// TwinCAT 3 PLC project PLC
// ProgramVersion: 3.1.4026.27
// CompilerDefines: VISU_USEPROPERTYINFO
// libraries:
//   Tc2_Standard, * (Beckhoff Automation GmbH)
//   Tc2_System, * (Beckhoff Automation GmbH)
//   Tc2_Utilities, * (Beckhoff Automation GmbH)
//   Tc3_DynamicMemory, * (Beckhoff Automation GmbH)
//   VisuDialogs, * (System)
//   VisuSymbols, 4.5.0.0 (System)
// project tree:
//   / GlobalTextList.TcGTLO, PlcTask.TcTTO, Visualization Manager.TcVMO (not stored)
//   POUs/ FB_Dynamic.TcPOU, MAIN.TcPOU, monoInstance.TcPOU, multiInstances.TcPOU
//   VISUs/ Visualization.TcVIS
// real-time tasks:
//   TASK PlcTask: cycle T#10ms, priority 20, ADS port 350

CONFIGURATION PLC
    RESOURCE PLC ON TwinCAT3
        TASK PlcTask(INTERVAL := T#10ms, PRIORITY := 20);
        PROGRAM MAIN WITH PlcTask : MAIN;
    END_RESOURCE
END_CONFIGURATION

// ---- POUs/MAIN.TcPOU
PROGRAM MAIN
VAR
(*
+--------------------------------------------------------------------------+
| PROGRAMME DE TEST - CREATION DYNAMIQUE (__NEW / __DELETE)                |
| TwinCAT 3 - IEC 61131-3 - Structured Text                                |
+--------------------------------------------------------------------------+
|                                                                          |
| Projet d'exemple TwinCAT 3 illustrant la creation et la destruction      |
| dynamiques d'instances de bloc fonction (FB) pendant l'execution du      |
| PLC, avec les operateurs __NEW et __DELETE.                              |
|                                                                          |
+--------------------------------------------------------------------------+
| monoInstance                                                             |
|   -> Creer / detruire une seule instance de FB_Dynamic                   |
+--------------------------------------------------------------------------+
| multiInstances                                                           |
|   -> Gerer un nombre dynamique d'instances (de 0 a cMaxInstances),       |
|      ajustable en ligne, avec suivi de la memoire du router              |
+--------------------------------------------------------------------------+
*)
END_VAR

//monoInstance();
multiInstances();

END_PROGRAM

// ---- POUs/multiInstances.TcPOU
PROGRAM multiInstances
VAR CONSTANT
    cMaxInstances : UINT := 1000;      // passer à 100, puis 1000 pour tester les limites
END_VAR
VAR
    // Tableau de pointeurs (aucune instance n'est créée statiquement)
    aFB            : ARRAY[1..cMaxInstances] OF POINTER TO FB_Dynamic;
    aResult        : ARRAY[1..cMaxInstances] OF INT;

    // Commande
    nTarget        : UINT := 10;     // nombre d'instances souhaité (modifiable en ligne)
    nMaxOpsPerCycle: UINT := 50;     // limite de __NEW/__DELETE par cycle
    nIncrease      : INT := 5;

    // Diagnostic
    nActive        : UINT;           // instances actuellement créées
    nNewFailed     : UDINT;          // nombre d'échecs de __NEW
    bAllocError    : BOOL;

    // Variables locales de travail
    i              : UINT;
    nOps           : UINT;

    // Surveillance du router (ton code existant)
    fbGetRouterStatusInfo : FB_GetRouterStatusInfo;
    TonGetRouterStatus    : TON;
    bError                : BOOL;
    nErrorID              : UDINT;
    stTcRouterStatusInfo  : Tc2_Utilities.ST_TcRouterStatusInfo;
	nUsage: REAL;
	bInc: BOOL;
	bDec: BOOL;
END_VAR

// --- 1. Ajustement du nombre d'instances vers nTarget ---
nTarget := LIMIT(0, nTarget, cMaxInstances);
nOps    := 0;

FOR i := 1 TO cMaxInstances DO
    IF nOps >= nMaxOpsPerCycle THEN
        EXIT;                              // on étale la charge sur plusieurs cycles
    END_IF

    IF i <= nTarget THEN
        // Instance souhaitée : on la crée si elle n'existe pas
        IF aFB[i] = 0 THEN
            aFB[i] := __NEW(FB_Dynamic);
            nOps := nOps + 1;
            IF aFB[i] = 0 THEN             // __NEW renvoie 0 si plus de mémoire
                nNewFailed  := nNewFailed + 1;
                bAllocError := TRUE;
                EXIT;
            END_IF
        END_IF
    ELSE
        // Instance en trop : on la détruit
        IF aFB[i] <> 0 THEN
            __DELETE(aFB[i]);
            aFB[i] := 0;                   // indispensable
            nOps := nOps + 1;
        END_IF
    END_IF
END_FOR

// --- 2. Appel cyclique des instances existantes ---
nActive := 0;
FOR i := 1 TO cMaxInstances DO
    IF aFB[i] <> 0 THEN
        aResult[i] := aFB[i]^.Increase(nCountStep := nIncrease);
        nActive    := nActive + 1;
    END_IF
END_FOR

// --- 3. Surveillance du router (inchangé) ---
fbGetRouterStatusInfo(
    sNetId   := '',
    bExecute := NOT TonGetRouterStatus.Q,
    tTimeout := DEFAULT_ADS_TIMEOUT,
    bBusy    => ,
    bError   => bError,
    nErrID   => nErrorID,
    info     => stTcRouterStatusInfo);

TonGetRouterStatus(IN := NOT fbGetRouterStatusInfo.bBusy, PT := T#1S);

IF stTcRouterStatusInfo.maxMem >0 THEN
nUsage:=(TO_REAL(stTcRouterStatusInfo.maxMem-stTcRouterStatusInfo.maxMemAvail)/TO_REAL(stTcRouterStatusInfo.maxMem))*100.0;
END_IF

IF bInc AND nTarget<cMaxInstances THEN
	nTarget:=nTarget+1;
	bInc:=FALSE;
END_IF

IF bDec  AND nTarget>1 THEN
	nTarget:=nTarget-1;
	bDec:=FALSE;
END_IF

END_PROGRAM

// ---- POUs/FB_Dynamic.TcPOU
{attribute 'enable_dynamic_creation'}
FUNCTION_BLOCK FB_Dynamic
VAR
    nCounts : INT;
END_VAR

METHOD Increase : INT
VAR_INPUT
	nCountStep :INT;
END_VAR
nCounts := nCounts + nCountStep;
Increase := nCounts;
END_METHOD

END_FUNCTION_BLOCK

// ---- POUs/monoInstance.TcPOU
PROGRAM monoInstance
VAR
	pFB       : POINTER TO FB_Dynamic;
    nResult   : INT;
    nIncrease : INT := 5;
    bNew      : BOOL := TRUE;
    bDelete   : BOOL;
	
	fbGetRouterStatusInfo:FB_GetRouterStatusInfo;
	TonGetRouterStatus:TON;
	bError: BOOL;
	nErrorID: UDINT;
	stTcRouterStatusInfo: Tc2_Utilities.ST_TcRouterStatusInfo;
END_VAR

IF bNew AND (pFB = 0) THEN
    pFB := __NEW(FB_Dynamic);
    bNew := FALSE;
END_IF

IF (pFB <> 0) THEN
    nResult := pFB^.Increase(nCountStep := nIncrease);
END_IF

IF bDelete THEN
    __DELETE(pFB);
    bDelete := FALSE;
END_IF


fbGetRouterStatusInfo(
	sNetId:= '', 
	bExecute:= NOT TonGetRouterStatus.Q, 
	tTimeout:= DEFAULT_ADS_TIMEOUT, 
	bBusy=> , 
	bError=> bError, 
	nErrID=> nErrorID, 
	info=> stTcRouterStatusInfo);

IF stTcRouterStatusInfo.maxMem >0 THEN
	TonGetRouterStatus(IN:= NOT fbGetRouterStatusInfo.bBusy, PT:=T#1S , Q=> , ET=> );
END_IF

END_PROGRAM

// ---- GlobalTextList.TcGTLO
TEXTLIST GlobalTextList
  77 = '+'
  247 = '-'
  9 = 'nb Instances %d'
  278 = 'nb Instances: %d'
  284 = 'nb Target: %d'
  238 = 'Usage : %.2f %'
  439 = 'Usage : %.2f%'
END_TEXTLIST

// ---- VISUs/Visualization.TcVIS
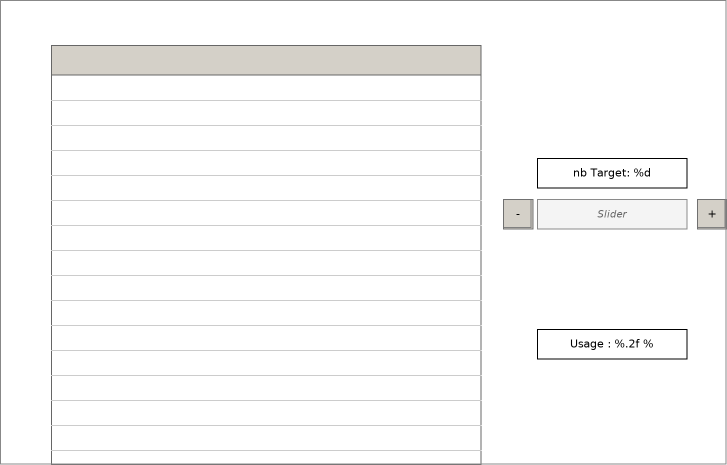
VISUALIZATION Visualization  // 727x465
    Table (51,45 430x420), data array: multiInstances.aFB
        p1128707560: multiInstances.cMaxInstances
        p3854506369: multiInstances.aFB[INDEX]^.nCounts
        p1014161805: MULTIINSTANCES.cMaxInstances - 1 + INT#1
    Rectangle (537,158 150x30), "nb Target: %d", text variable: multiInstances.nTarget
        OnMouseClick: write the text variable via Default, min 1, max multiInstances.cMaxInstances
    Rectangle (537,329 150x30), "Usage : %.2f %", text variable: multiInstances.nUsage
    Slider (537,199 150x30), variable: multiInstances.nTarget, scale 1..100
    Button (697,199 30x30), "+"
        OnMouseClick: toggle multiInstances.bInc
    Button (503,199 30x30), "-"
        OnMouseClick: toggle multiInstances.bDec
END_VISUALIZATION
